// Palpeur Keyence GT2, type 31 (docs/03 § 6.2), mode signaux : S1 AI valeur. Le mode réseau (P1 = 1) n'est pas
// encore écrit : la configuration est refusée.
// Hypothèse : la valeur brute de l'entrée analogique est en micromètres (1 = 0,001 mm), comme la sortie
// analogique du GT2 réglée sur ±32 mm. À confirmer avec le câblage réel.
FUNCTION_BLOCK FB_KeyenceGT2 EXTENDS FB_ObjectBase
VAR
    _fValue : LREAL;                // mm, après remise à zéro
    _fRaw : LREAL;                  // mm, avant remise à zéro
    _fZero : LREAL;
    _bOutOfRange : BOOL;
    _fStabMs : LREAL;
    _nWanted : INT;
    _nTaken : INT;
    _fSum : LREAL;
    _fSimValue : LREAL;
END_VAR
VAR PERSISTENT
    _fZeroKept : LREAL;             // remise à zéro gardée après une coupure
END_VAR

METHOD PROTECTED _OnConfigure : BOOL
IF _bNewObject THEN _fZeroKept := 0; END_IF
_fZero := _fZeroKept;
_fSimValue := _refCfg.aParam[2];
_OnConfigure := _refCfg.aParam[1] = 0 AND F_SignalValid(_refCfg.aSignal[1], E_SignalKind.AI);
END_METHOD

METHOD PROTECTED _OnStart : E_ActStatus
VAR_INPUT
    nAction : UINT;
END_VAR
CASE nAction OF
    GVL_Catalog.KeyenceGT2_Mesurer:
        _nWanted := LIMIT(1, LREAL_TO_INT(_ParamReal(1, _refCfg.aParam[5])), 1000);
        _nTaken := 0;
        _fSum := 0;
        _fStabMs := 0;
        _OnStart := E_ActStatus.Busy;
    GVL_Catalog.KeyenceGT2_RemiseAZero:
        _fZero := _fRaw;
        _fZeroKept := _fZero;
        _OnStart := E_ActStatus.Done;
    GVL_Catalog.KeyenceGT2_LireValeurCourante:
        _SetResult(1, _fValue);
        _OnStart := E_ActStatus.Done;
ELSE
    _OnStart := E_ActStatus.Error;
END_CASE
END_METHOD

METHOD PROTECTED _OnCycle : E_ActStatus
VAR_INPUT
    nAction : UINT;
END_VAR
VAR
    fMean : LREAL;
    fHigh : LREAL;
    fLow : LREAL;
END_VAR
_OnCycle := E_ActStatus.Busy;
IF _bOutOfRange THEN
    _Fail(GVL_Catalog.KeyenceGT2_Err100, 0);
    _OnCycle := E_ActStatus.Error;
    RETURN;
END_IF
// Stabilisation P6, puis un échantillon par cycle
_fStabMs := _fStabMs + F_CycleMs();
IF _fStabMs < MAX(0.0, _refCfg.aParam[6]) THEN RETURN; END_IF
_fSum := _fSum + _fValue;
_nTaken := _nTaken + 1;
IF _nTaken < _nWanted THEN RETURN; END_IF
fMean := _fSum / INT_TO_LREAL(_nTaken);
fHigh := _refCfg.aParam[2] + ABS(_refCfg.aParam[3]);
fLow := _refCfg.aParam[2] - ABS(_refCfg.aParam[4]);
_SetResult(1, fMean);
IF fMean > fHigh THEN
    _SetJudgement(2, E_Judgement.High);
ELSIF fMean < fLow THEN
    _SetJudgement(2, E_Judgement.Low);
ELSE
    _SetJudgement(2, E_Judgement.Ok);
END_IF
_OnCycle := E_ActStatus.Done;
END_METHOD

METHOD PROTECTED _ReadHw
VAR
    nRaw : INT;
END_VAR
nRaw := F_ReadAI(_refCfg.aSignal[1]);
_bOutOfRange := nRaw = 32767 OR nRaw = -32768;
_fRaw := INT_TO_LREAL(nRaw) * 0.001;
_fValue := _fRaw - _fZero;
END_METHOD

// Simulation : valeur de référence P2 avec un bruit de ±10 % de la tolérance haute (docs/03 § 6.2)
METHOD PROTECTED _Simulate
_fRaw := _fSimValue + (F_SimRandom() - 0.5) * 0.2 * ABS(_refCfg.aParam[3]) + _fZero;
IF _Forced(1) THEN _fRaw := _ForcedValue(1) + _fZero; END_IF       // valeur forcée en mm
_bOutOfRange := FALSE;
_fValue := _fRaw - _fZero;
END_METHOD

METHOD PROTECTED _Publish
_stStatus.aValue[1] := _fValue;
END_METHOD

END_FUNCTION_BLOCK

(* stored: Version 1.1.0.1, ProductVersion 3.1.4024.12
   POU FB_KeyenceGT2: Id {039a6318-8c79-503d-b91a-1c6412a9aa03}, SpecialFunc None
   Method _OnConfigure: Id {8ab515f2-db78-52cc-a133-1da6a0957e55}
   Method _OnStart: Id {1006cf16-337d-5b6c-a2a6-b28394001753}
   Method _OnCycle: Id {e05a3722-907e-5b6a-b15d-61c5afb5e1ad}
   Method _ReadHw: Id {54563a8a-3abf-5887-9a07-0fc636c50bd0}
   Method _Simulate: Id {3c6fd347-d852-5bdf-9b99-f48926886bf7}
   Method _Publish: Id {22a19cac-e864-5c1a-a3c5-69ec0226d8f8} *)
